Fanuc KAREL source: KO00111.KL

PROGRAM KO00111
%NOLOCKGROUP
VAR
  A: REAL
  B: ARRAY[2] OF SHORT
  OUT: INTEGER
BEGIN
  A = 1
  B[1] = 2
  OUT = ATAN2(A, B[1])
END KO00111
